(* IEC 61131-3 sources: TetherPLC/tools/oracle/corpus, 21 files *)

(* ---- conv_case.st ---- *)
PROGRAM Demo
VAR
    t1 AT %QD0  : DINT;
    ro AT %QD4  : DINT;
    m1 AT %QD8  : DINT;
    m2 AT %QD12 : DINT;
    u1 AT %QD16 : UDINT;
END_VAR
t1 := TRUNC(-3.9);
ro := ROUND(2.5);
m1 := MUX(1, 10, 20, 30);
m2 := MUX(2, 10, 20, 30);
u1 := DINT_TO_UDINT(7);
END_PROGRAM

(* ---- ctd_case.st ---- *)
PROGRAM CtdCase
VAR
    dn   AT %IX0.0 : BOOL;
    load AT %IX0.1 : BOOL;
    done AT %QX0.0 : BOOL;
    ctd1 : CTD;
END_VAR
ctd1(CD := dn, LD := load, PV := 3);
done := ctd1.QD;
END_PROGRAM

(* ---- ctu_case.st ---- *)
PROGRAM CtuCase
VAR
    pulse AT %IX0.0 : BOOL;
    reset AT %IX0.1 : BOOL;
    done AT %QX0.0 : BOOL;
    ctu1 : CTU;
    last_cv : INT;
END_VAR
ctu1(CU := pulse, R := reset, PV := 3);
done := ctu1.QU;
last_cv := ctu1.CV;
END_PROGRAM

(* ---- divzero_case.st ---- *)
PROGRAM Demo
VAR
    d AT %ID0 : DINT;
    e AT %ID4 : DINT;
    out AT %QD0 : DINT;
    out2 AT %QD4 : DINT;
END_VAR
out := 100 / d;
out2 := 103 MOD e;
END_PROGRAM

(* ---- fn_case.st ---- *)
PROGRAM Demo
VAR
    s     : STRING[16];
    t     : STRING[16];
    c     : STRING[32];
    w     : WSTRING[16];
    wc    : WSTRING[32];
    n1 AT %QD0    : DINT;
    flags AT %QD4 : DINT;
END_VAR
s := 'abc';
t := 'xyz';
c := CONCAT(s, t);
w := "aä";
wc := CONCAT(w, w);
n1 := LEN(c);
flags := 0;
IF c = 'abcxyz' THEN
    flags := flags + 1;
END_IF
IF LEN(wc) = 4 THEN
    flags := flags + 2;
END_IF
IF wc = "aäaä" THEN
    flags := flags + 4;
END_IF
END_PROGRAM

(* ---- ovf_case.st ---- *)
PROGRAM OvfCase
VAR
    a AT %ID0 : DINT;
    b AT %ID4 : DINT;
    s AT %IW8 : INT;
    n AT %IW10 : INT;
    out AT %QD0 : DINT;
    out2 AT %QW4 : INT;
    out3 AT %QW6 : INT;
    out4 AT %QD8 : DINT;
END_VAR
out := a + b;
out2 := s * 1000;
out3 := -n;
out4 := a - b;
END_PROGRAM

(* ---- ovf_div.st ---- *)
PROGRAM OvfDiv
VAR
    a AT %IL0 : LINT;
    b AT %IL8 : LINT;
    out AT %QL0 : LINT;
    out2 AT %QL8 : LINT;
END_VAR
out := a / b;
out2 := a + b;
END_PROGRAM

(* ---- ref_case.st ---- *)
PROGRAM Demo
VAR
    x   : DINT := 42;
    r   : REFERENCE TO DINT;
    out AT %QD0 : DINT;
    ok  AT %QD4 : DINT;
END_VAR
r REF= x;
out := r;
ok := 0;
IF ISVALIDREF(r) THEN
    ok := ok + 1;
END_IF
IF r^ = 42 THEN
    ok := ok + 2;
END_IF
IF r = 42 THEN
    ok := ok + 4;
END_IF
END_PROGRAM

(* ---- rng_case.st ---- *)
PROGRAM RngCase
VAR
    d AT %ID0 : DINT;
    r AT %IL8 : LREAL;
    u AT %ID16 : UDINT;
    out AT %QD0 : DINT;
    out2 AT %QD4 : DINT;
    out3 AT %QD8 : DINT;
    out4 AT %QD12 : DINT;
END_VAR
out := DINT_TO_INT(d);
out2 := LREAL_TO_DINT(r);
out3 := DINT_TO_UINT(d);
out4 := UDINT_TO_DINT(u);
END_PROGRAM

(* ---- rtrig_case.st ---- *)
PROGRAM RTrigCase
VAR
    sig  AT %IX0.0 : BOOL;
    rise AT %QX0.0 : BOOL;
    fall AT %QX0.1 : BOOL;
    rt1  : R_TRIG;
    ft1  : F_TRIG;
END_VAR
rt1(CLK := sig);
ft1(CLK := sig);
rise := rt1.Q;
fall := ft1.Q;
END_PROGRAM

(* ---- scalar_fn.st ---- *)
PROGRAM Demo
VAR
    a AT %QD0  : DINT;
    b AT %QD4  : DINT;
    c AT %QD8  : DINT;
    d AT %QD12 : DINT;
    e AT %QD16 : DINT;
    f AT %QD20 : DINT;
END_VAR
a := ABS(-5);
b := MIN(3, 7);
c := MAX(3, 7);
d := SEL(FALSE, 11, 22);
e := LIMIT(10, 42, 20);
f := ABS(4 - 9);
END_PROGRAM

(* ---- sh_active.st ---- *)
PROGRAM ShActive
VAR
    cnt : DINT;
    out_cnt AT %QD0 : DINT;
END_VAR
cnt := cnt + 1;
out_cnt := cnt;
END_PROGRAM

(* ---- sh_cand_b.st ---- *)
PROGRAM ShActive
VAR
    cnt : DINT;
    out_cnt AT %QD0 : DINT;
END_VAR
cnt := cnt + 1;
out_cnt := 3 * cnt;
END_PROGRAM

(* ---- sh_cand_c.st ---- *)
PROGRAM ShActive
VAR
    cnt : DINT;
    out_cnt AT %QD0 : DINT;
END_VAR
cnt := cnt + 1;
out_cnt := 4 * cnt;
END_PROGRAM

(* ---- sh_candidate.st ---- *)
PROGRAM ShActive
VAR
    cnt : DINT;
    out_cnt AT %QD0 : DINT;
END_VAR
cnt := cnt + 1;
out_cnt := 2 * cnt;
END_PROGRAM

(* ---- srrs_case.st ---- *)
PROGRAM SrRsCase
VAR
    a   AT %IX0.0 : BOOL;
    b   AT %IX0.1 : BOOL;
    qsr AT %QX0.0 : BOOL;
    qrs AT %QX0.1 : BOOL;
    sr1 : SR;
    rs1 : RS;
END_VAR
sr1(S1 := a, R := b);
rs1(S := a, R1 := b);
qsr := sr1.Q1;
qrs := rs1.Q1;
END_PROGRAM

(* ---- str_case.st ---- *)
PROGRAM Demo
VAR
    a  : STRING[16];
    b  : STRING[16];
    eq1 AT %QX0.0 : BOOL;
    eq2 AT %QX0.1 : BOOL;
    eq3 AT %QX0.2 : BOOL;
    eq4 AT %QX0.3 : BOOL;
    eq5 AT %QX0.4 : BOOL;
END_VAR
a := 'abc';
b := 'abd';
eq1 := (a = b);
eq2 := (a = 'abc');
eq3 := (a <> b);
eq4 := ('ab' = 'ab');
eq5 := ('ab' = 'abc');
END_PROGRAM

(* ---- strfn_case.st ---- *)
PROGRAM Demo
VAR
    s  : STRING[16];
    t  : STRING[16];
    ok AT %QD0 : DINT;
    n1 AT %QD4 : DINT;
END_VAR
s := 'abcdef';
t := 'XY';
ok := 0;
IF LEFT(s, 3) = 'abc' THEN
    ok := ok + 1;
END_IF
IF RIGHT(s, 3) = 'def' THEN
    ok := ok + 2;
END_IF
IF MID(s, 2, 3) = 'cd' THEN
    ok := ok + 4;
END_IF
IF INSERT(s, t, 4) = 'abcXYdef' THEN
    ok := ok + 8;
END_IF
IF DELETE(s, 2, 3) = 'abef' THEN
    ok := ok + 16;
END_IF
IF REPLACE(s, t, 2, 3) = 'abXYef' THEN
    ok := ok + 32;
END_IF
n1 := FIND(s, 'cd');
END_PROGRAM

(* ---- tof_case.st ---- *)
PROGRAM TofCase
VAR
    sig  AT %IX0.0 : BOOL;
    outp AT %QX0.0 : BOOL;
    tof1 : TOF;
END_VAR
tof1(IN := sig, PT := T#500ms);
outp := tof1.Q;
END_PROGRAM

(* ---- ton_case.st ---- *)
PROGRAM TonCase
VAR
    start_in AT %IX0.0 : BOOL;
    lamp AT %QX0.0 : BOOL;
    ton1 : TON;
    et_seen : TIME;
END_VAR
ton1(IN := start_in, PT := T#500ms);
lamp := ton1.Q;
et_seen := ton1.ET;
END_PROGRAM

(* ---- wstr_case.st ---- *)
PROGRAM Demo
VAR
    w  : WSTRING[16];
    w2 : WSTRING[16];
    eq1 AT %QX0.0 : BOOL;
    eq2 AT %QX0.1 : BOOL;
    eq3 AT %QX0.2 : BOOL;
END_VAR
w := "abc";
w2 := "abd";
eq1 := (w = w2);
eq2 := (w = "abc");
eq3 := (w <> w2);
END_PROGRAM
